(* IEC 61131-3 sources: plc-ci-toolkit/ci/tests/samples/sa_probe_src/src/POUs/PRG_Main, 2 files *)

(* ---- PRG_Main.decl.st ---- *)
// Назначение: главная программа примера. Обрабатывает однократные команды HMI
//             (квитирование, сброс через интерфейс I_Resettable), вызывает FB_Example
//             и публикует состояние для HMI. Обмен с HMI — через stCmd и stSts.
// Автор:      kr0nsch
// Версия:     0.1.0
// Документ:   docs/ARCHITECTURE.md, раздел «Пример в src/»
PROGRAM PRG_Main
VAR
    fbPump : FB_Example;            // насос подкачки: регулирование по уровню
    itfResettable : I_Resettable;   // сброс через интерфейс — одинаково для любых ФБ с I_Resettable
    stCmd : ST_ExampleCmd;          // команды HMI/SCADA
    stSts : ST_ExampleSts;          // состояние для HMI/SCADA
    rLevel_pct : REAL;              // уровень, % — привязать к входу модуля или задать онлайн
    xLevelValid : BOOL;             // достоверность уровня (в проекте — результат проверки NE 43)
    xPumpOn : BOOL;                 // команда на пускатель насоса — привязать к выходу модуля
    fbSaBad : FB_SaBad;
    fbSaSkip : FB_SaSkip;
    xTmp : BOOL;
END_VAR

(* ---- PRG_Main.impl.st ---- *)
// 1. Однократные команды HMI выполняем до вызова ФБ, чтобы выход в этом же цикле
//    отражал результат; после выполнения команду сбрасывает ПЛК.
IF stCmd.xAck THEN
    stCmd.xAck := FALSE;
    fbPump.Acknowledge();
END_IF

IF stCmd.xReset THEN
    stCmd.xReset := FALSE;
    itfResettable := fbPump;
    itfResettable.Reset();
END_IF

// 2. Регулирование
fbPump(eMode := stCmd.eMode,
       rValue_pct := rLevel_pct,
       xValueValid := xLevelValid,
       rSetpoint_pct := stCmd.rSetpoint_pct,
       xManualOn := stCmd.xManualOn,
       xOut => xPumpOn);

// 3. Состояние для HMI
stSts.eMode := stCmd.eMode;
stSts.xOut := xPumpOn;
stSts.xFault := fbPump.xFault;
stSts.rSetpointUsed_pct := fbPump.rSetpointUsed_pct;
stSts.udiCount := fbPump.Count;

// зонд статанализа
fbSaBad(iMode := 1, rIn := 1.5);
xTmp := fbSaBad.Check() AND F_SaTemp(xIn := TRUE);
GVL_SaProbe.diShared := 5;
GVL_SaProbe.xOutBad := xTmp;
GVL_SaProbe.wOverlapA := 1;
GVL_SaProbe.bOverlapB := 2;
fbSaSkip(xIn := xTmp);
